Universal Robots URScript: T002_mistralai_Mistral-Large-3-675B-Instruct-2512-NVFP4_edit_perf_rep1.urscript

# Task: T002 — Linear weld path — fenced mode (Optimized for cycle time)
# Robot: ur5e
# Operating mode: fenced | Max TCP speed: 0.500 m/s

def task_T002():
  TCP_SPEED_CAP = 0.500
  def safe_movel(pose, a, v, r):
    if (v > TCP_SPEED_CAP):
      popup("TCP speed cap exceeded", error=True)
      halt
    end
    movel(pose, a=a, v=v, r=r)
  end

  # [0] Verify E-Stop clear before weld sequence
  if (get_digital_in(0) == True):
    popup("E-Stop active — aborting program.", error=True)
    halt
  end

  # [1] Go to home position (increased speed)
  movej([0.0000, -1.5708, 1.5708, -1.5708, -1.5708, 0.0000], a=2.0000, v=1.2000)

  # [2] Approach above weld start (increased speed)
  safe_movel(p[0.450000, 0.000000, 0.350000, 0.0000, 3.1416, 0.0000], 1.5000, 0.4000, 0.0100)

  # [3] Descend to weld start position (increased acceleration)
  safe_movel(p[0.450000, 0.000000, 0.200000, 0.0000, 3.1416, 0.0000], 1.0000, 0.1500, 0.0010)

  # [4] Gas pre-flow ON (parallel with motion)
  set_digital_out(1, True)

  # [5] Gas stabilization delay (reduced)
  sleep(0.3000)

  # [6] Arc ON — welding start
  set_digital_out(0, True)
  set_analog_out(0, 0.400)
  set_analog_out(1, 0.333)

  # [7] Weld seam — 300mm linear path (optimized speed)
  safe_movel(p[0.450000, 0.300000, 0.200000, 0.0000, 3.1416, 0.0000], 0.5000, 0.0500, 0.0)

  # [8] Arc OFF — welding end
  set_digital_out(0, False)
  set_analog_out(0, 0.0)
  set_analog_out(1, 0.0)

  # [9] Post-weld gas flow (reduced)
  sleep(0.5000)

  # [10] Gas flow OFF
  set_digital_out(1, False)

  # [11] Retract above weld end (increased speed)
  safe_movel(p[0.450000, 0.300000, 0.350000, 0.0000, 3.1416, 0.0000], 1.5000, 0.4000, 0.0100)

  # [12] Return to home (increased speed)
  movej([0.0000, -1.5708, 1.5708, -1.5708, -1.5708, 0.0000], a=2.0000, v=1.2000)
end

# Entry point
task_T002()
